FUNCTION_BLOCK T_SafeMon_Tests EXTENDS TcUnit.FB_TestSuite
VAR
    // Test_AutomaticRestartWhenGuardClosed
    group_1 : T_SafeGroup;
    fb_1 : T_SafeMon(group := group_1);
    // Test_SecureInputBypassesGuard
    group_2 : T_SafeGroup;
    fb_2 : T_SafeMon(group := group_2);
    // Test_ManualFunctionTestRequiresGuardOpenedOnce
    group_3 : T_SafeGroup;
    fb_3 : T_SafeMon(group := group_3) := (Parameters := (ManualFunctionTest := TRUE));
    // Test_EdmFaultWithoutManualRestartStaysSafe
    group_4 : T_SafeGroup;
    fb_4 : T_SafeMon(group := group_4);
    // Test_NoMonInConnectedIsRefused
    group_5 : T_SafeGroup;
    fb_5 : T_SafeMon(group := group_5);
    // Test_ResetTimeNotMultipleOfTenIsRefused
    group_6 : T_SafeGroup;
    fb_6 : T_SafeMon(group := group_6) := (Parameters := (Edm1ResetTime := T#15MS));
END_VAR

Test_AutomaticRestartWhenGuardClosed();
Test_SecureInputBypassesGuard();
Test_ManualFunctionTestRequiresGuardOpenedOnce();
Test_EdmFaultWithoutManualRestartStaysSafe();
Test_NoMonInConnectedIsRefused();
Test_ResetTimeNotMultipleOfTenIsRefused();

METHOD PRIVATE Test_AutomaticRestartWhenGuardClosed
TcUnit.TEST(__POUNAME());
// act: Restart not connected -> automatic restart; guard open
group_1(Run := TRUE);
fb_1(MonIn1 := FALSE);
group_1(Run := TRUE);
fb_1(MonIn1 := FALSE);
// assert
AssertEquals_BOOL(Expected := FALSE, Actual := fb_1.MonOut, Message := 'output off with guard open');
group_1(Run := TRUE);
fb_1(MonIn1 := TRUE);
AssertEquals_BOOL(Expected := TRUE, Actual := fb_1.MonOut, Message := 'automatic restart with guard closed');
AssertEquals_BYTE(Expected := TO_BYTE(E_SafeMonState.Run), Actual := fb_1.State, Message := 'state RUN');
TEST_FINISHED_NAMED(__POUNAME());
END_METHOD

METHOD PRIVATE Test_EdmFaultWithoutManualRestartStaysSafe
TcUnit.TEST(__POUNAME());
// act: EDM1 connected and FALSE, no Restart connected
group_4(Run := TRUE);
fb_4(EDM1 := FALSE, MonIn1 := TRUE);
group_4(Run := TRUE);
fb_4(EDM1 := FALSE, MonIn1 := TRUE);
// assert
AssertEquals_BOOL(Expected := FALSE, Actual := fb_4.Error, Message := 'no EDM error without manual restart');
AssertEquals_BYTE(Expected := TO_BYTE(E_SafeMonState.Safe), Actual := fb_4.State, Message := 'FB remains SAFE');
TEST_FINISHED_NAMED(__POUNAME());
END_METHOD

METHOD PRIVATE Test_ManualFunctionTestRequiresGuardOpenedOnce
TcUnit.TEST(__POUNAME());
// arrange: Restart connected (manual restart), guard closed from the start
group_3(Run := TRUE);
fb_3(Restart := FALSE, MonIn1 := TRUE);
AssertEquals_BYTE(Expected := TO_BYTE(E_SafeMonState.FuncTest), Actual := fb_3.State, Message := 'state FUNCTEST after start');
// act: restart without testing the guard
group_3(Run := TRUE);
fb_3(Restart := TRUE, MonIn1 := TRUE);
group_3(Run := TRUE);
fb_3(Restart := FALSE, MonIn1 := TRUE);
AssertEquals_BOOL(Expected := FALSE, Actual := fb_3.MonOut, Message := 'restart ignored before the function test');
// act: open and close the guard, then restart
group_3(Run := TRUE);
fb_3(Restart := FALSE, MonIn1 := FALSE);
group_3(Run := TRUE);
fb_3(Restart := FALSE, MonIn1 := TRUE);
group_3(Run := TRUE);
fb_3(Restart := TRUE, MonIn1 := TRUE);
group_3(Run := TRUE);
fb_3(Restart := FALSE, MonIn1 := TRUE);
AssertEquals_BOOL(Expected := TRUE, Actual := fb_3.MonOut, Message := 'output on after function test and restart');
TEST_FINISHED_NAMED(__POUNAME());
END_METHOD

METHOD PRIVATE Test_SecureInputBypassesGuard
TcUnit.TEST(__POUNAME());
// act: guard open, bypass active
group_2(Run := TRUE);
fb_2(MonIn1 := FALSE, Secure1 := TRUE);
group_2(Run := TRUE);
fb_2(MonIn1 := FALSE, Secure1 := TRUE);
// assert
AssertEquals_BOOL(Expected := TRUE, Actual := fb_2.MonOut, Message := 'guard ignored while Secure is 1');
group_2(Run := TRUE);
fb_2(MonIn1 := FALSE, Secure1 := FALSE);
AssertEquals_BOOL(Expected := FALSE, Actual := fb_2.MonOut, Message := 'guard monitored again when Secure is 0');
TEST_FINISHED_NAMED(__POUNAME());
END_METHOD

METHOD PRIVATE Test_NoMonInConnectedIsRefused
TcUnit.TEST(__POUNAME());
// arrange / act: only the Secure pair is connected, which the Safety Editor refuses
group_5(Run := TRUE);
fb_5(Secure1 := TRUE);
group_5(Run := TRUE);
fb_5(Secure1 := TRUE);
// assert
AssertEquals_BOOL(Expected := TRUE, Actual := fb_5.Error, Message := 'configuration error reported');
AssertEquals_BYTE(Expected := TO_BYTE(E_SafeFbState.Error), Actual := fb_5.State, Message := 'state ERROR');
AssertEquals_WORD(Expected := WORD#16#8000, Actual := fb_5.Diag, Message := 'diag bit 15 configuration refused');
AssertEquals_BOOL(Expected := FALSE, Actual := fb_5.MonOut, Message := 'MonOut stays at its safe value');
AssertEquals_BOOL(Expected := TRUE, Actual := group_5.FbErr, Message := 'the group sees an FB error');
// act: ErrAck 0 -> 1 -> 0 does not clear a configuration error
group_5(Run := TRUE, ErrAck := TRUE);
fb_5(Secure1 := TRUE);
group_5(Run := TRUE, ErrAck := TRUE);
fb_5(Secure1 := TRUE);
group_5(Run := TRUE, ErrAck := FALSE);
fb_5(Secure1 := TRUE);
AssertEquals_BOOL(Expected := TRUE, Actual := fb_5.Error, Message := 'error not acknowledged');
AssertEquals_WORD(Expected := WORD#16#8000, Actual := fb_5.Diag, Message := 'diag bit 15 kept');
TEST_FINISHED_NAMED(__POUNAME());
END_METHOD

METHOD PRIVATE Test_ResetTimeNotMultipleOfTenIsRefused
TcUnit.TEST(__POUNAME());
// arrange / act: Edm1ResetTime is 15 ms, which the Safety Editor refuses
group_6(Run := TRUE);
fb_6(EDM1 := TRUE, MonIn1 := TRUE);
group_6(Run := TRUE);
fb_6(EDM1 := TRUE, MonIn1 := TRUE);
// assert
AssertEquals_BOOL(Expected := TRUE, Actual := fb_6.Error, Message := 'configuration error reported');
AssertEquals_BYTE(Expected := TO_BYTE(E_SafeFbState.Error), Actual := fb_6.State, Message := 'state ERROR');
AssertEquals_WORD(Expected := WORD#16#8000, Actual := fb_6.Diag, Message := 'diag bit 15 configuration refused');
AssertEquals_BOOL(Expected := FALSE, Actual := fb_6.MonOut, Message := 'MonOut stays at its safe value');
AssertEquals_BOOL(Expected := TRUE, Actual := group_6.FbErr, Message := 'the group sees an FB error');
// act: ErrAck 0 -> 1 -> 0 does not clear a configuration error
group_6(Run := TRUE, ErrAck := TRUE);
fb_6(EDM1 := TRUE, MonIn1 := TRUE);
group_6(Run := TRUE, ErrAck := TRUE);
fb_6(EDM1 := TRUE, MonIn1 := TRUE);
group_6(Run := TRUE, ErrAck := FALSE);
fb_6(EDM1 := TRUE, MonIn1 := TRUE);
AssertEquals_BOOL(Expected := TRUE, Actual := fb_6.Error, Message := 'error not acknowledged');
AssertEquals_WORD(Expected := WORD#16#8000, Actual := fb_6.Diag, Message := 'diag bit 15 kept');
TEST_FINISHED_NAMED(__POUNAME());
END_METHOD

END_FUNCTION_BLOCK

(* stored: Version 1.1.0.1
   POU T_SafeMon_Tests: Id {f06f20f6-051a-5cea-acd9-faf06a097146}, SpecialFunc None
   Method Test_AutomaticRestartWhenGuardClosed: Id {7f7524c0-8cb8-53ff-8d3a-e39d36e3ba99}
   Method Test_EdmFaultWithoutManualRestartStaysSafe: Id {35b5b4d2-365a-5ee9-8d58-df81715760f5}
   Method Test_ManualFunctionTestRequiresGuardOpenedOnce: Id {cf8948bc-d028-54a1-9163-5666b9b64e98}
   Method Test_SecureInputBypassesGuard: Id {76d3bf1a-d2bf-5feb-a26a-e6cd0e1dd4d6}
   Method Test_NoMonInConnectedIsRefused: Id {0e51c03a-757d-4eeb-8e11-d119df2c4072}
   Method Test_ResetTimeNotMultipleOfTenIsRefused: Id {e61b8ec8-e7bb-4d34-aa76-4458974c248a} *)
